FUNCTION_BLOCK FB_EL3356ChannelDiagnosis
VAR_INPUT
	stChannelState				:ST_EL3356ChannelState;
END_VAR
VAR_OUTPUT
	bChannelOK					:BOOL;
	bCalibrationInProgress			:BOOL;
END_VAR
VAR

END_VAR


(* General Channel Status *)
IF stChannelState.bOverrange = 0
    AND stChannelState.bError = 0
    AND stChannelState.bSyncError = 0
THEN
	bChannelOK := TRUE;
ELSE
	bChannelOK := FALSE;
END_IF

bCalibrationInProgress := stChannelState.bCalibrationInProgress;

END_FUNCTION_BLOCK

(* stored: Version 1.1.0.1, ProductVersion 3.1.4024.15
   POU FB_EL3356ChannelDiagnosis: Id {15a6fda7-b4df-475b-b964-d0c172334a21}, SpecialFunc None *)
